Fanuc KAREL source: KT00713.KL

PROGRAM KT00713
%NOLOCKGROUP
VAR
  S1: STRING[80]
  S2: STRING[80]
  OUT: INTEGER
BEGIN
  S1 = 'A'
  S2 = 'B'
  S1 = 'A'
  S2 = 'B'
  OUT = ARRAY_LEN(S1)
END KT00713
